(*
SPDX-FileCopyrightText: © 2026 Oleksandr Tiutyk <trofimich@gmail.com>
SPDX-License-Identifier: MIT
License: https://opensource.org/license/mit
*)

(*!
<summary>Orders UDINT values described by generic descriptors.</summary>
<description>
Non-null addresses must reference live UDINT storage. TypeClass and Size are not validated and no numeric
conversion is performed. Two null addresses compare equal; one null address sorts before a non-null address.
Descriptors are passed by value; payload remains borrowed and is not modified, cloned, released or retained.
IsMemoryOwner does not affect comparison.
</description>
*)

FUNCTION_BLOCK UDIntComparer EXTENDS TOF_Core.Object IMPLEMENTS TOF_Core.IComparer
VAR_STAT
	//! <summary>Class name shared by all instances of this function block.</summary>
	{attribute 'hide'} 
	_ClassName : STRING := __POUNAME();
END_VAR

{attribute 'monitoring' := 'call'}
PROPERTY ClassName : REFERENCE TO STRING
GET
ClassName REF= _ClassName;
END_GET
END_PROPERTY

(*!
<summary>Compares the first operand with the second using this ordering strategy.</summary>
<description>
Non-null addresses must reference live UDINT storage. TypeClass and Size are not validated and no numeric
conversion is performed. Two null addresses compare equal; one null address sorts before a non-null address.
Descriptors are passed by value; payload remains borrowed and is not modified, cloned, released or retained.
IsMemoryOwner does not affect comparison. Descendants cannot replace this standard ordering; implement
IComparer separately for a different ordering strategy.
</description>
*)
//!<param name="first">First descriptor; referenced storage is borrowed for the call.</param>
//!<param name="second">Second descriptor; referenced storage is borrowed for the call.</param>
{attribute "object_name" := "Compare"}
METHOD FINAL Compare : TOF_Core.COMPARISON_RESULT
VAR_INPUT
	first : TOF_Core.GENERIC_VALUE;
	second : TOF_Core.GENERIC_VALUE;
END_VAR
VAR
	leftPointer : POINTER TO UDINT; 
	rightPointer : POINTER TO UDINT; 
END_VAR
IF first.Address = 0 AND_THEN second.Address = 0 THEN
	Compare := TOF_Core.COMPARISON_RESULT.FIRST_EQUAL_TO_SECOND;
	RETURN;
END_IF

IF first.Address = 0 THEN
	Compare := TOF_Core.COMPARISON_RESULT.FIRST_LESS_THAN_SECOND;
	RETURN;	
END_IF

IF second.Address = 0 THEN
	Compare := TOF_Core.COMPARISON_RESULT.FIRST_GREATER_THAN_SECOND;
	RETURN;	
END_IF

leftPointer := first.Address;
rightPointer := second.Address;

IF leftPointer^ < rightPointer^ THEN
	Compare := TOF_Core.COMPARISON_RESULT.FIRST_LESS_THAN_SECOND;
ELSIF leftPointer^ > rightPointer^ THEN
	Compare := TOF_Core.COMPARISON_RESULT.FIRST_GREATER_THAN_SECOND;
ELSE
	Compare := TOF_Core.COMPARISON_RESULT.FIRST_EQUAL_TO_SECOND;	
END_IF
END_METHOD

{attribute 'monitoring' := 'call'}
PROPERTY NamespaceName : REFERENCE TO STRING
GET
NamespaceName REF= CurrentNamespace.Name;
END_GET
END_PROPERTY

{attribute 'monitoring' := 'call'}
PROPERTY SelfSize : ULINT
GET
SelfSize := XSIZEOF(THIS^);
END_GET
END_PROPERTY

END_FUNCTION_BLOCK

(* stored: Version 1.1.0.1
   POU UDIntComparer: Id {0ae69507-8f7d-48b2-9728-39bafe49b500}, SpecialFunc None
   Property ClassName: Id {07094e12-1afe-4df0-a577-00770f59e141}
   Get Get: Id {0c2a89c1-020f-4e90-992a-e9c92ab6a9e5}
   Method Compare: Id {189176fb-e2b7-4029-9aa3-41432925664d}
   Property NamespaceName: Id {57216ce7-1543-4b07-9467-ab7ebf55ccbd}
   Get Get: Id {cb2a1877-6c14-4ea9-b444-415e77728225}
   Property SelfSize: Id {afdf47e5-4760-49ff-a8d5-f1ebd7c5fa1e}
   Get Get: Id {a08f4458-d60c-4849-b78d-6c3956be1f49} *)
